RoboDK station: pick and place sencillo.rdk

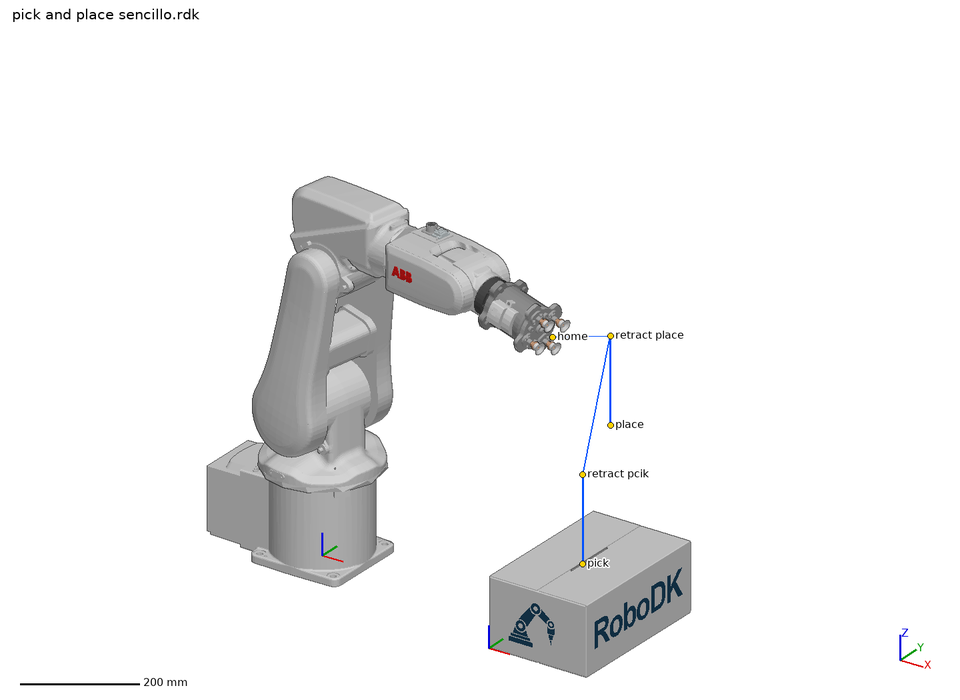
[picture v0: the station drawn from its stored meshes, robots at their saved joint values, targets as dots, program paths as lines]
Station pick and place sencillo (saved by RoboDK 5.5.0). Poses are relative to the parent item; angles as X-Y-Z fixed-axis rotations.
  - frame ABB IRB 120-3/0.6 Base at (0, 0, 0) mm
    - robot ABB IRB 120-3/0.6: 6 axes, payload 3 kg, reach 580 mm, repeatability 0.01 mm, weight 25 kg
        modified DH rows (alpha deg, a mm, theta deg, d mm): 0, 0, 0, 290; -90, 0, -90, 0; 0, 270, 0, 0; -90, 70, 0, 302; 90, 0, 0, 0; -90, 0, 180, 72
        joint limits [-165, -110, -90, -160, -120, -400] to [165, 110, 70, 160, 120, 400]; home [0, 0, 0, 0, 0, 0]; saved at [-10, 10, -10, 0, 10, -20]
      - tool SMC ZXP7A01-ZP20U-X1 Vacuum Gripper, TCP at (0, 0, 125) mm, size 88 x 106.8 x 127.9 mm
  - frame Frame 2 at (430, -130, 0) mm
    - object Box 12x7in (Closed) at (0, 0, 0) mm, size 199 x 305.1 x 133.7 mm, geometry from Box-12x7in-Closed.sld
    - target pick (Cartesian target) at (100.37, 130, 132.62) mm, rotated rx 180 ry 0 rz 180 deg; joints [0, 60.43, -29.803, 0, 59.373, 0] of ABB IRB 120-3/0.6
    - target retract pcik (Cartesian target) at (100.37, 130, 297.62) mm, rotated rx 180 ry 0 rz -180 deg; joints [0, 56.627, -54.002, 0, 87.375, 0] of ABB IRB 120-3/0.6
    - target retract place (Cartesian target) at (-164.81, 589.32, 297.67) mm, rotated rx 180 ry 0.01 rz -120 deg; joints [60, 56.62, -54, 0, 87.37, 0] of ABB IRB 120-3/0.6
    - target place (Cartesian target) at (-164.82, 589.31, 132.61) mm, rotated rx 180 ry 0 rz -120 deg; joints [60, 60.43, -29.8, 0, 59.37, 0] of ABB IRB 120-3/0.6
    - target home (Cartesian target) at (104.64, 35.73, 591.69) mm, rotated rx -117.27 ry 67.73 rz -125.51 deg; joints [-10, 10, -10, 0, 10, -20] of ABB IRB 120-3/0.6
  - program pickandplace (11 instructions, listed below)
  - program Reset (1 instructions, listed below)
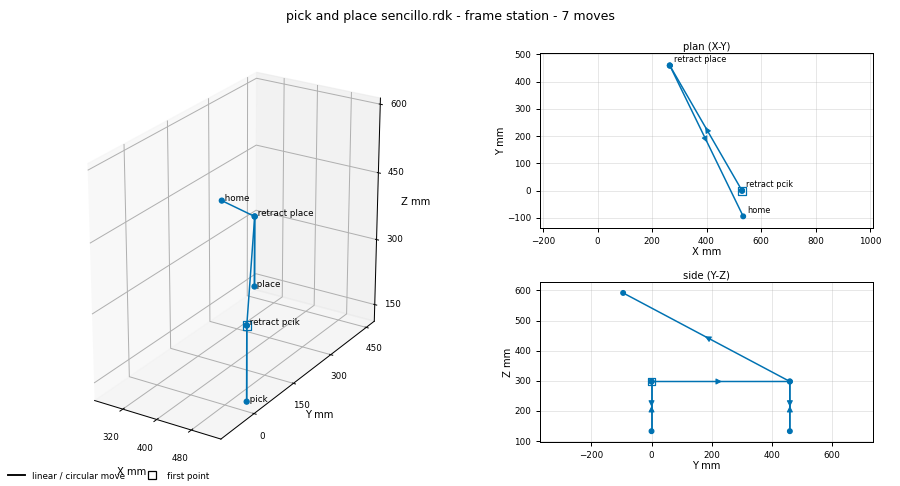
[picture p0: tool path of pick and place sencillo.rdk in frame station, 7 of 7 moves have a stored position in this frame; points joined in program order, loops and branches not executed]

--- program pickandplace (robot ABB IRB 120-3/0.6) ---
  Est. Ref.: Frame 2
  Est. herr: SMC ZXP7A01-ZP20U-X1 Vacuum Gripper
  MoveJ (retract pcik)
  MoveL (pick)
  Adjuntar a SMC ZXP7A01-ZP20U-X1 Vacuum Gripper
  MoveL (retract pcik)
  MoveL (retract place)
  MoveL (place)
  Separar de SMC ZXP7A01-ZP20U-X1 Vacuum Gripper
  MoveL (retract place)
  MoveL (home)

--- program Reset (robot ABB IRB 120-3/0.6) ---
  Reemplazar Box 12x7in (Closed)
